// TIA Portal V21 export
// export: Created 2026-11-08T21:48:03.8206839Z, ExportSetting WithDefaults, DisplayName Totally Integrated Automation Portal, DisplayVersion V21 Update 3, DisplayName STEP 7 Professional, DisplayVersion V21 Update 3, DisplayName STEP 7 Safety, DisplayVersion V21, DisplayName Tech WebApplication, DisplayVersion V21, DisplayName WinCC Basic/Comfort/Advanced, DisplayVersion V21 Update 3, DisplayName WinCC Unified, DisplayVersion V21 Update 3
DATA_BLOCK "FB_Khp_DB"   // DB7
// stored: AutoNumber true, DBAccessibleFromOPCUA true, DBAccessibleFromWebserver true, InstanceOfName FB_Khp, InstanceOfType FB
"FB_Khp"
   // VAR_INPUT
   //    inp : Int;
   // END_VAR
   // VAR_OUTPUT
   //    outp : Bool;
   // END_VAR
   // VAR
   //    st : Real;
   //    tmr { S7_SetPoint := 'True'} : TON_TIME;
   // END_VAR
BEGIN
END_DATA_BLOCK
